Fanuc KAREL source: kc00048.KL

-- PROVISIONAL review KL for V1013-1; original PC SHA256 1ecf577b4125397c36d3297236fc15ba37000ac7adc997e418f5aef2fa81ec2c
-- Incomplete behavior may be omitted. Consult companion uncertainty JSON. Do not deploy.
PROGRAM KC00048
%NOLOCKGROUP
BEGIN
  -- UNRESOLVED_PC offsets 5-35; opcodes 27,22,22,1C,22,27,9D,31
  -- UNRESOLVED_PC offsets 40-44; opcodes 7F
END KC00048
